// TIA Portal V21 export
// export: Created 2026-11-02T09:43:47.7393727Z, ExportSetting WithDefaults, DisplayName Totally Integrated Automation Portal, DisplayVersion V21 Update 3, DisplayName TIA Portal Test Suite Advanced, DisplayVersion V21 Update 1, DisplayName SINAMICS Startdrive Advanced, DisplayVersion V21 Update 1, DisplayName SINAMICS Startdrive G130, G150, S120, S150, G200, G210, G210C, G210X, G220, S200, S210, S220, Innomotics MVD, DisplayVersion V21 Update 1, DisplayName SINAMICS Startdrive G110M, G120, G120C, G120D, G120P, G115D, DisplayVersion V21 Update 1, DisplayName STEP 7 Professional, DisplayVersion V21 Update 3, DisplayName STEP 7 Safety, DisplayVersion V21, DisplayName Tech WebApplication, DisplayVersion V21, DisplayName WinCC Basic/Comfort/Advanced, DisplayVersion V21 Update 3, DisplayName WinCC Professional, DisplayVersion V21 Update 3, DisplayName WinCC Unified, DisplayVersion V21 Update 3
FUNCTION_BLOCK "Tgp_TON_LAD"   // FB2, LAD
{ S7_Optimized_Access := 'TRUE' }
VERSION : 0.1
// stored: AutoNumber true, IsIECCheckEnabled false, IsRetainMemResEnabled false, MemoryReserve 100, SetENOAutomatically false, UDAEnableTagReadback false
   VAR_INPUT
      Enable : Bool;
      Preset : Time;
   END_VAR
   VAR_OUTPUT
      Done : Bool;
      Elapsed : Time;
   END_VAR
   VAR
      Storage { S7_SetPoint := 'True'} : TON_TIME;
   END_VAR
BEGIN

REGION Network 1
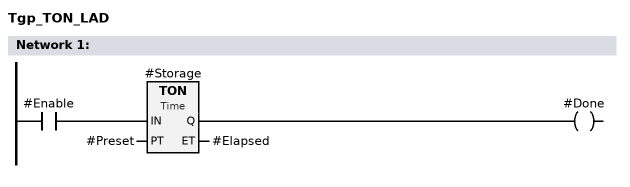
   RUNG wire#powerrail
      Contact( #Enable )
      { S7_Templates := "time_type := Time" } #Storage.TON(pt := #Preset, et => #Elapsed)
      Coil( #Done )
   END_RUNG
   // the same network as SCL:
   #Storage(IN := #Enable, PT := #Preset, ET => #Elapsed);   // TON
   #Done := #Storage.Q;
END_REGION
END_FUNCTION_BLOCK
